FUNCTION FC 1 : VOID
BEGIN
NETWORK
      A X 0.0
END_FUNCTION
